// TIA Portal V15.1 export
// export: Created 2026-11-02T18:55:11.1503167Z, ExportSetting WithDefaults, DisplayName Totally Integrated Automation Portal, DisplayVersion V15.1, DisplayName TIA Portal Openness, DisplayVersion V15.1, DisplayName STEP 7 Professional, DisplayVersion V15.1, DisplayName WinCC Professional, DisplayVersion V15.1
DATA_BLOCK "Scrubber_DB"   // DB5
{ S7_Optimized_Access := 'TRUE' }
VERSION : 0.1
// stored: AutoNumber false, InstanceOfName Scrubber, InstanceOfType FB
"Scrubber"
   // VAR_INPUT
   //    PSH : Bool;
   //    LSH : Bool;
   //    LSHH : Bool;
   //    EStopOK : Bool;
   //    ResetPulse : Bool;
   //    FirstScan : Bool;
   //    TDrnOn : Time;
   //    TDrnOff : Time;
   //    TDrnMax : Time;
   // END_VAR
   // VAR_OUTPUT
   //    Tripped : Bool;
   //    FlareTrip : Bool;
   //    ValvesNormal : Bool;
   //    FlareCmd : Bool;
   //    DrainCmd : Bool;
   //    SuctionCmd : Bool;
   //    F_DrainTO : Bool;
   //    F_LshFault : Bool;
   //    Alm_PSH : Bool;
   //    Alm_LSH : Bool;
   //    Alm_LSHH : Bool;
   //    Cause_EStop : Bool;
   //    Cause_PSH : Bool;
   //    Cause_LSHH : Bool;
   //    Cause_PwrUp : Bool;
   //    FirstOut : Int;
   // END_VAR
   // VAR
   //    LevelHigh : Bool;
   //    DrnDemand : Bool;
   //    T_DrnOn : TON_TIME;
   //    T_DrnOff : TON_TIME;
   //    T_DrnMax : TON_TIME;
   //    T_LshFlt : TON_TIME;
   // END_VAR
BEGIN
END_DATA_BLOCK
